Staubli VAL3: utData.dtx

public num nVal
public bool bStatus
